(* IEC 61131-3 sources: rules_plc/examples/simple_2, 2 files *)

(* ---- mathlib.st ---- *)
FUNCTION_BLOCK st_add
    VAR_INPUT
        a : DINT;
        b : DINT;
    END_VAR
    VAR_OUTPUT
        out: DINT;
    END_VAR
    VAR
        call_count : DINT;
    END_VAR
    call_count := call_count + 1;
    out := a + b;
END_FUNCTION_BLOCK

FUNCTION st_double : DINT
    VAR_INPUT
        x : DINT;
    END_VAR
    st_double := x * 2;
END_FUNCTION

(* ---- doubler_app.st ---- *)
{external}
FUNCTION puts : DINT
    VAR_INPUT {ref}
        text : STRING;
    END_VAR
END_FUNCTION

PROGRAM doubler_app
    VAR
        result : DINT;
    END_VAR
    result := st_double(21);
    puts('doubled value computed$N');
END_PROGRAM
